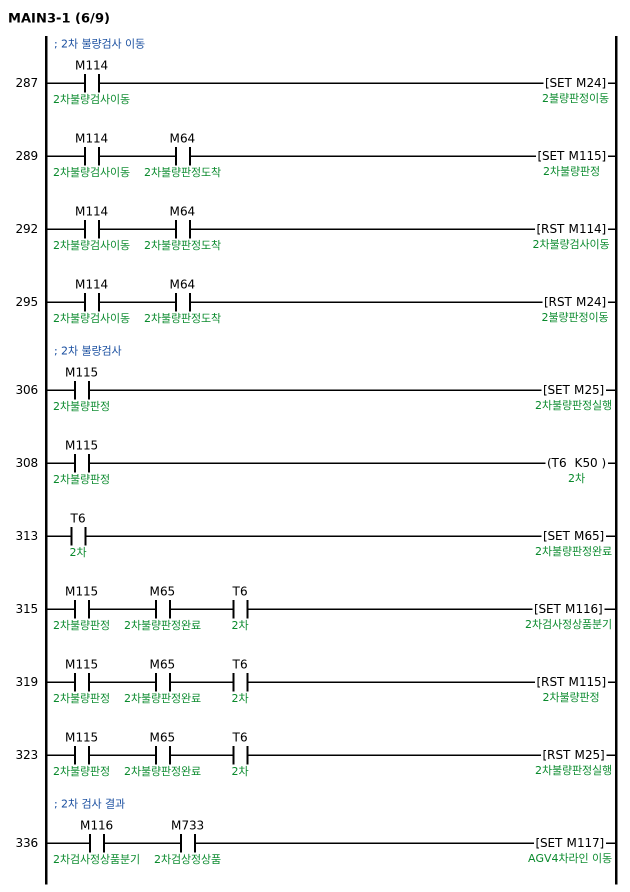
; 2차 불량검사 이동
287   LD      M114  ; 2차불량검사이동
      SET     M24  ; 2불량판정이동
289   LD      M114  ; 2차불량검사이동
      AND     M64  ; 2차불량판정도착
      SET     M115  ; 2차불량판정
292   LD      M114  ; 2차불량검사이동
      AND     M64  ; 2차불량판정도착
      RST     M114  ; 2차불량검사이동
295   LD      M114  ; 2차불량검사이동
      AND     M64  ; 2차불량판정도착
      RST     M24  ; 2불량판정이동
; 2차 불량검사
306   LD      M115  ; 2차불량판정
      SET     M25  ; 2차불량판정실행
308   LD      M115  ; 2차불량판정
      OUT     T6 K50  ; 2차
313   LD      T6  ; 2차
      SET     M65  ; 2차불량판정완료
315   LD      M115  ; 2차불량판정
      AND     M65  ; 2차불량판정완료
      AND     T6  ; 2차
      SET     M116  ; 2차검사정상품분기
319   LD      M115  ; 2차불량판정
      AND     M65  ; 2차불량판정완료
      AND     T6  ; 2차
      RST     M115  ; 2차불량판정
323   LD      M115  ; 2차불량판정
      AND     M65  ; 2차불량판정완료
      AND     T6  ; 2차
      RST     M25  ; 2차불량판정실행
; 2차 검사 결과
336   LD      M116  ; 2차검사정상품분기
      AND     M733  ; 2차검상정상품
      SET     M117  ; AGV4차라인 이동
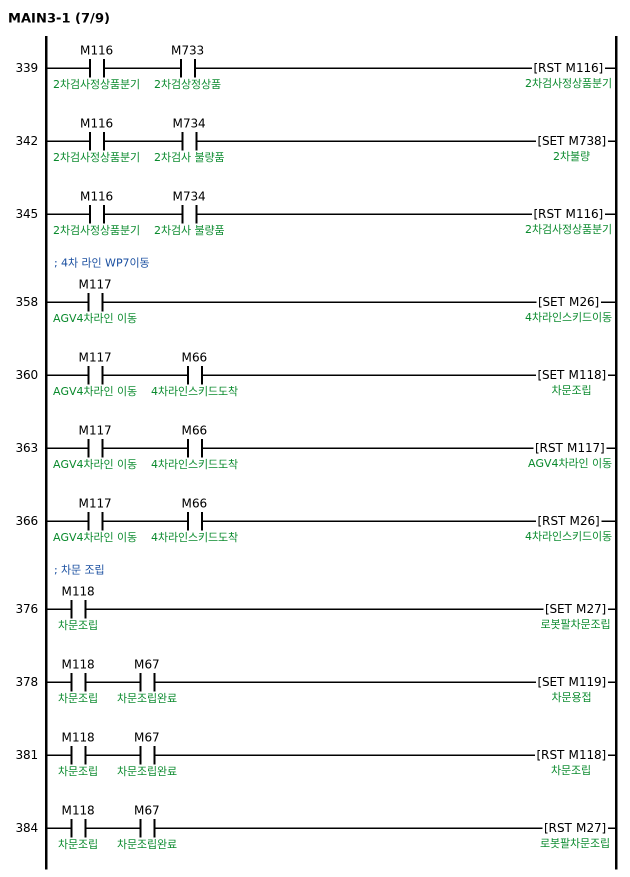
339   LD      M116  ; 2차검사정상품분기
      AND     M733  ; 2차검상정상품
      RST     M116  ; 2차검사정상품분기
342   LD      M116  ; 2차검사정상품분기
      AND     M734  ; 2차검사 불량품
      SET     M738  ; 2차불량
345   LD      M116  ; 2차검사정상품분기
      AND     M734  ; 2차검사 불량품
      RST     M116  ; 2차검사정상품분기
; 4차 라인 WP7이동
358   LD      M117  ; AGV4차라인 이동
      SET     M26  ; 4차라인스키드이동
360   LD      M117  ; AGV4차라인 이동
      AND     M66  ; 4차라인스키드도착
      SET     M118  ; 차문조립
363   LD      M117  ; AGV4차라인 이동
      AND     M66  ; 4차라인스키드도착
      RST     M117  ; AGV4차라인 이동
366   LD      M117  ; AGV4차라인 이동
      AND     M66  ; 4차라인스키드도착
      RST     M26  ; 4차라인스키드이동
; 차문 조립
376   LD      M118  ; 차문조립
      SET     M27  ; 로봇팔차문조립
378   LD      M118  ; 차문조립
      AND     M67  ; 차문조립완료
      SET     M119  ; 차문용접
381   LD      M118  ; 차문조립
      AND     M67  ; 차문조립완료
      RST     M118  ; 차문조립
384   LD      M118  ; 차문조립
      AND     M67  ; 차문조립완료
      RST     M27  ; 로봇팔차문조립
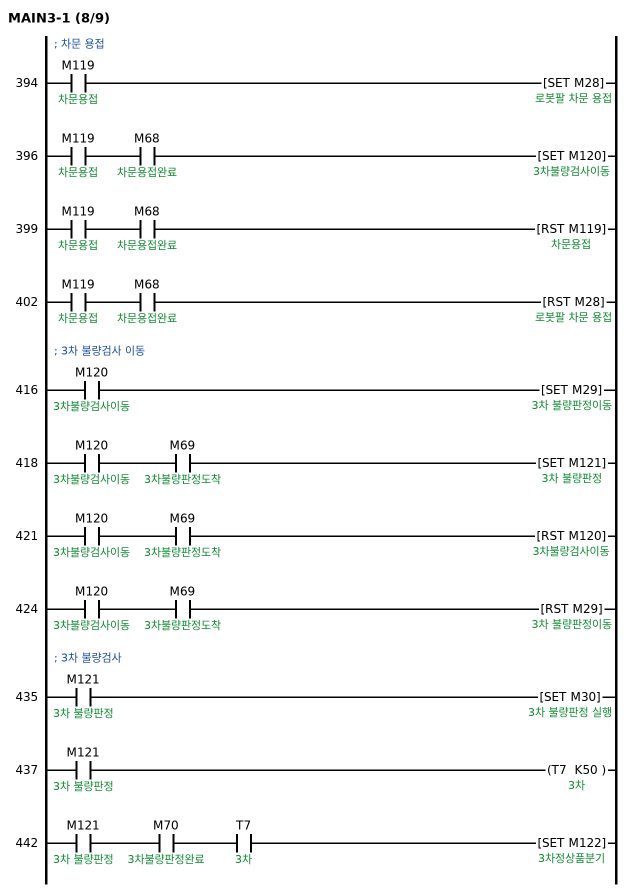
; 차문 용접
394   LD      M119  ; 차문용접
      SET     M28  ; 로봇팔 차문 용접
396   LD      M119  ; 차문용접
      AND     M68  ; 차문용접완료
      SET     M120  ; 3차불량검사이동
399   LD      M119  ; 차문용접
      AND     M68  ; 차문용접완료
      RST     M119  ; 차문용접
402   LD      M119  ; 차문용접
      AND     M68  ; 차문용접완료
      RST     M28  ; 로봇팔 차문 용접
; 3차 불량검사 이동
416   LD      M120  ; 3차불량검사이동
      SET     M29  ; 3차 불량판정이동
418   LD      M120  ; 3차불량검사이동
      AND     M69  ; 3차불량판정도착
      SET     M121  ; 3차 불량판정
421   LD      M120  ; 3차불량검사이동
      AND     M69  ; 3차불량판정도착
      RST     M120  ; 3차불량검사이동
424   LD      M120  ; 3차불량검사이동
      AND     M69  ; 3차불량판정도착
      RST     M29  ; 3차 불량판정이동
; 3차 불량검사
435   LD      M121  ; 3차 불량판정
      SET     M30  ; 3차 불량판정 실행
437   LD      M121  ; 3차 불량판정
      OUT     T7 K50  ; 3차
442   LD      M121  ; 3차 불량판정
      AND     M70  ; 3차불량판정완료
      AND     T7  ; 3차
      SET     M122  ; 3차정상품분기
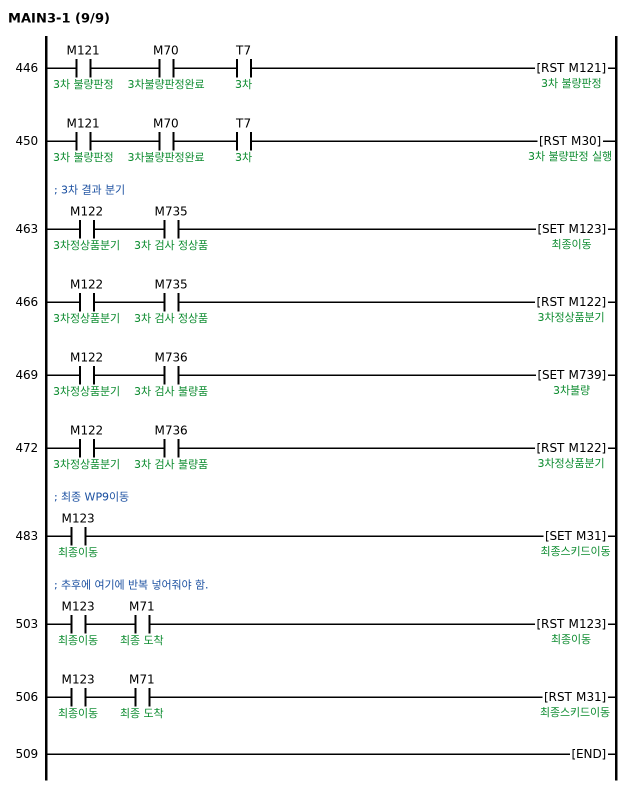
446   LD      M121  ; 3차 불량판정
      AND     M70  ; 3차불량판정완료
      AND     T7  ; 3차
      RST     M121  ; 3차 불량판정
450   LD      M121  ; 3차 불량판정
      AND     M70  ; 3차불량판정완료
      AND     T7  ; 3차
      RST     M30  ; 3차 불량판정 실행
; 3차 결과 분기
463   LD      M122  ; 3차정상품분기
      AND     M735  ; 3차 검사 정상품
      SET     M123  ; 최종이동
466   LD      M122  ; 3차정상품분기
      AND     M735  ; 3차 검사 정상품
      RST     M122  ; 3차정상품분기
469   LD      M122  ; 3차정상품분기
      AND     M736  ; 3차 검사 불량품
      SET     M739  ; 3차불량
472   LD      M122  ; 3차정상품분기
      AND     M736  ; 3차 검사 불량품
      RST     M122  ; 3차정상품분기
; 최종 WP9이동
483   LD      M123  ; 최종이동
      SET     M31  ; 최종스키드이동
; 추후에 여기에 반복 넣어줘야 함.
503   LD      M123  ; 최종이동
      AND     M71  ; 최종 도착
      RST     M123  ; 최종이동
506   LD      M123  ; 최종이동
      AND     M71  ; 최종 도착
      RST     M31  ; 최종스키드이동
509   END
END_PROGRAM

PROGRAM MAIN2-1
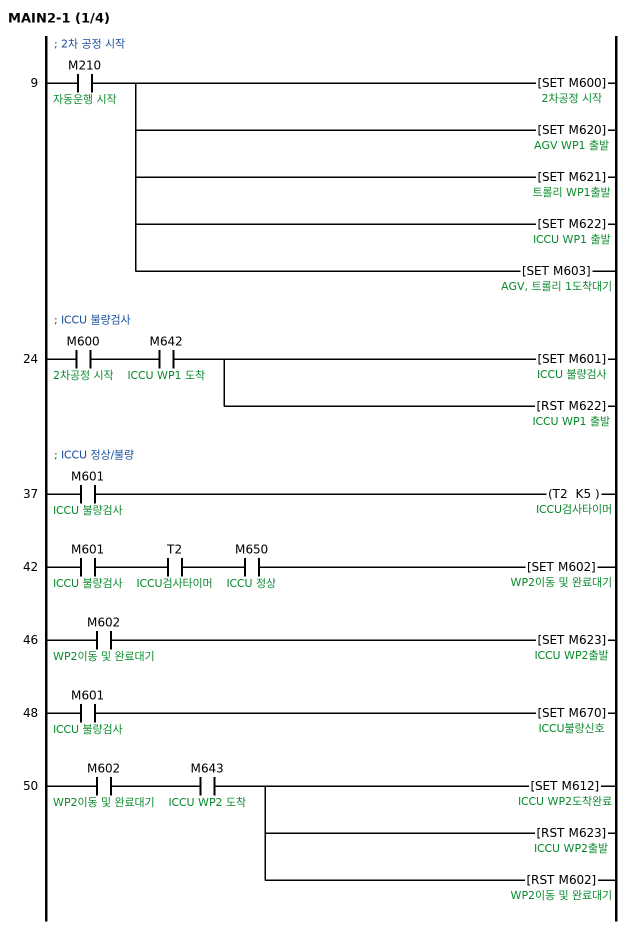
; 2차 공정 시작
9     LD      M210  ; 자동운행 시작
      SET     M600  ; 2차공정 시작
      SET     M620  ; AGV WP1 출발
      SET     M621  ; 트롤리 WP1출발
      SET     M622  ; ICCU WP1 출발
      SET     M603  ; AGV, 트롤리 1도착대기
; ICCU 불량검사
24    LD      M600  ; 2차공정 시작
      AND     M642  ; ICCU WP1 도착
      SET     M601  ; ICCU 불량검사
      RST     M622  ; ICCU WP1 출발
; ICCU 정상/불량
37    LD      M601  ; ICCU 불량검사
      OUT     T2 K5  ; ICCU검사타이머
42    LD      M601  ; ICCU 불량검사
      AND     T2  ; ICCU검사타이머
      AND     M650  ; ICCU 정상
      SET     M602  ; WP2이동 및 완료대기
46    LD      M602  ; WP2이동 및 완료대기
      SET     M623  ; ICCU WP2출발
48    LD      M601  ; ICCU 불량검사
      SET     M670  ; ICCU불량신호
50    LD      M602  ; WP2이동 및 완료대기
      AND     M643  ; ICCU WP2 도착
      SET     M612  ; ICCU WP2도착완료
      RST     M623  ; ICCU WP2출발
      RST     M602  ; WP2이동 및 완료대기
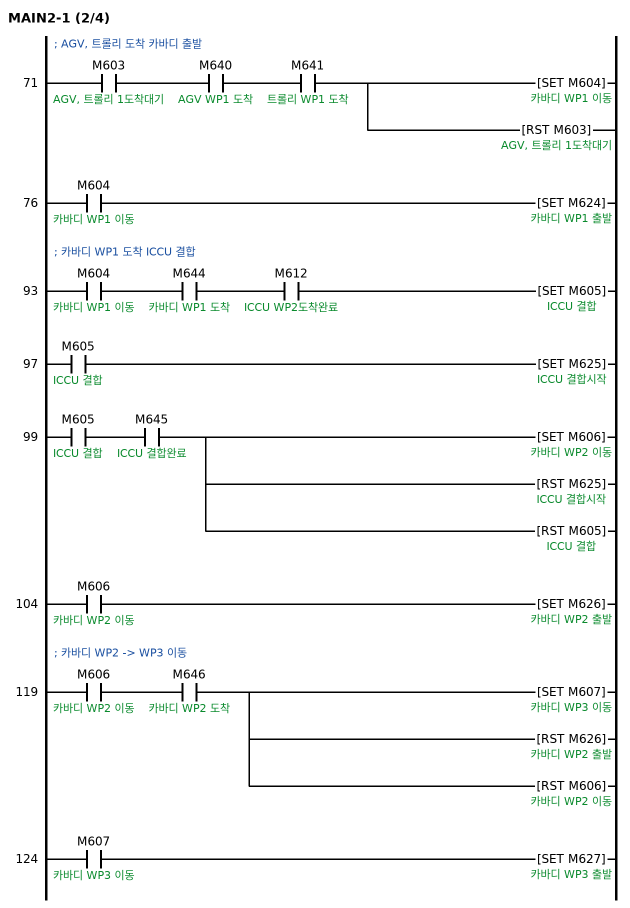
; AGV, 트롤리 도착 카바디 출발
71    LD      M603  ; AGV, 트롤리 1도착대기
      AND     M640  ; AGV WP1 도착
      AND     M641  ; 트롤리 WP1 도착
      SET     M604  ; 카바디 WP1 이동
      RST     M603  ; AGV, 트롤리 1도착대기
76    LD      M604  ; 카바디 WP1 이동
      SET     M624  ; 카바디 WP1 출발
; 카바디 WP1 도착 ICCU 결합
93    LD      M604  ; 카바디 WP1 이동
      AND     M644  ; 카바디 WP1 도착
      AND     M612  ; ICCU WP2도착완료
      SET     M605  ; ICCU 결합
97    LD      M605  ; ICCU 결합
      SET     M625  ; ICCU 결합시작
99    LD      M605  ; ICCU 결합
      AND     M645  ; ICCU 결합완료
      SET     M606  ; 카바디 WP2 이동
      RST     M625  ; ICCU 결합시작
      RST     M605  ; ICCU 결합
104   LD      M606  ; 카바디 WP2 이동
      SET     M626  ; 카바디 WP2 출발
; 카바디 WP2 -> WP3 이동
119   LD      M606  ; 카바디 WP2 이동
      AND     M646  ; 카바디 WP2 도착
      SET     M607  ; 카바디 WP3 이동
      RST     M626  ; 카바디 WP2 출발
      RST     M606  ; 카바디 WP2 이동
124   LD      M607  ; 카바디 WP3 이동
      SET     M627  ; 카바디 WP3 출발
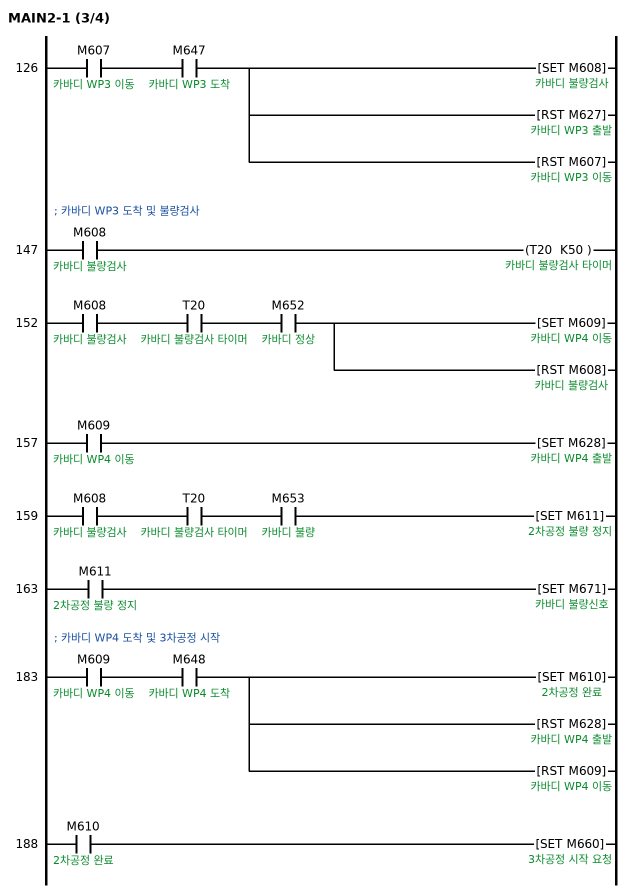
126   LD      M607  ; 카바디 WP3 이동
      AND     M647  ; 카바디 WP3 도착
      SET     M608  ; 카바디 불량검사
      RST     M627  ; 카바디 WP3 출발
      RST     M607  ; 카바디 WP3 이동
; 카바디 WP3 도착 및 불량검사
147   LD      M608  ; 카바디 불량검사
      OUT     T20 K50  ; 카바디 불량검사 타이머
152   LD      M608  ; 카바디 불량검사
      AND     T20  ; 카바디 불량검사 타이머
      AND     M652  ; 카바디 정상
      SET     M609  ; 카바디 WP4 이동
      RST     M608  ; 카바디 불량검사
157   LD      M609  ; 카바디 WP4 이동
      SET     M628  ; 카바디 WP4 출발
159   LD      M608  ; 카바디 불량검사
      AND     T20  ; 카바디 불량검사 타이머
      AND     M653  ; 카바디 불량
      SET     M611  ; 2차공정 불량 정지
163   LD      M611  ; 2차공정 불량 정지
      SET     M671  ; 카바디 불량신호
; 카바디 WP4 도착 및 3차공정 시작
183   LD      M609  ; 카바디 WP4 이동
      AND     M648  ; 카바디 WP4 도착
      SET     M610  ; 2차공정 완료
      RST     M628  ; 카바디 WP4 출발
      RST     M609  ; 카바디 WP4 이동
188   LD      M610  ; 2차공정 완료
      SET     M660  ; 3차공정 시작 요청
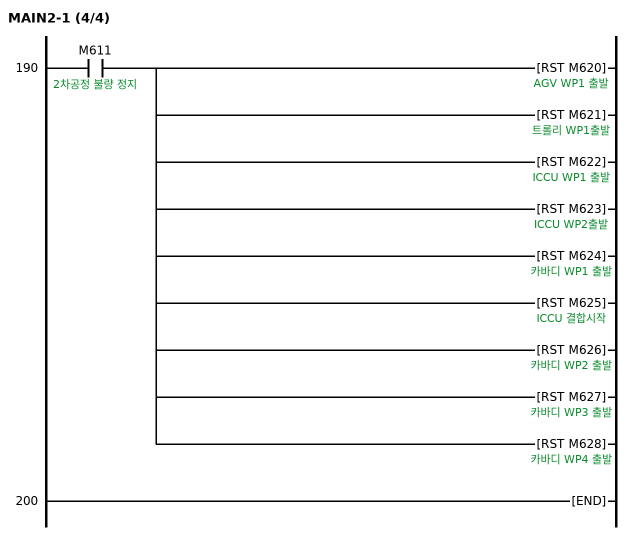
190   LD      M611  ; 2차공정 불량 정지
      RST     M620  ; AGV WP1 출발
      RST     M621  ; 트롤리 WP1출발
      RST     M622  ; ICCU WP1 출발
      RST     M623  ; ICCU WP2출발
      RST     M624  ; 카바디 WP1 출발
      RST     M625  ; ICCU 결합시작
      RST     M626  ; 카바디 WP2 출발
      RST     M627  ; 카바디 WP3 출발
      RST     M628  ; 카바디 WP4 출발
200   END
END_PROGRAM

PROGRAM MAIN2-2
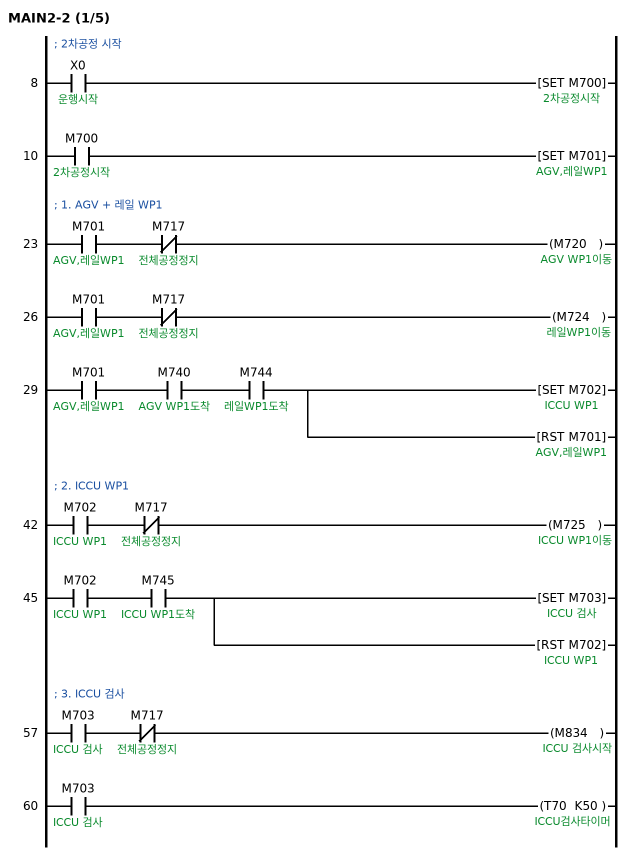
; 2차공정 시작
8     LD      X0  ; 운행시작
      SET     M700  ; 2차공정시작
10    LD      M700  ; 2차공정시작
      SET     M701  ; AGV,레일WP1
; 1. AGV + 레일 WP1
23    LD      M701  ; AGV,레일WP1
      ANI     M717  ; 전체공정정지
      OUT     M720  ; AGV WP1이동
26    LD      M701  ; AGV,레일WP1
      ANI     M717  ; 전체공정정지
      OUT     M724  ; 레일WP1이동
29    LD      M701  ; AGV,레일WP1
      AND     M740  ; AGV WP1도착
      AND     M744  ; 레일WP1도착
      SET     M702  ; ICCU WP1
      RST     M701  ; AGV,레일WP1
; 2. ICCU WP1
42    LD      M702  ; ICCU WP1
      ANI     M717  ; 전체공정정지
      OUT     M725  ; ICCU WP1이동
45    LD      M702  ; ICCU WP1
      AND     M745  ; ICCU WP1도착
      SET     M703  ; ICCU 검사
      RST     M702  ; ICCU WP1
; 3. ICCU 검사
57    LD      M703  ; ICCU 검사
      ANI     M717  ; 전체공정정지
      OUT     M834  ; ICCU 검사시작
60    LD      M703  ; ICCU 검사
      OUT     T70 K50  ; ICCU검사타이머
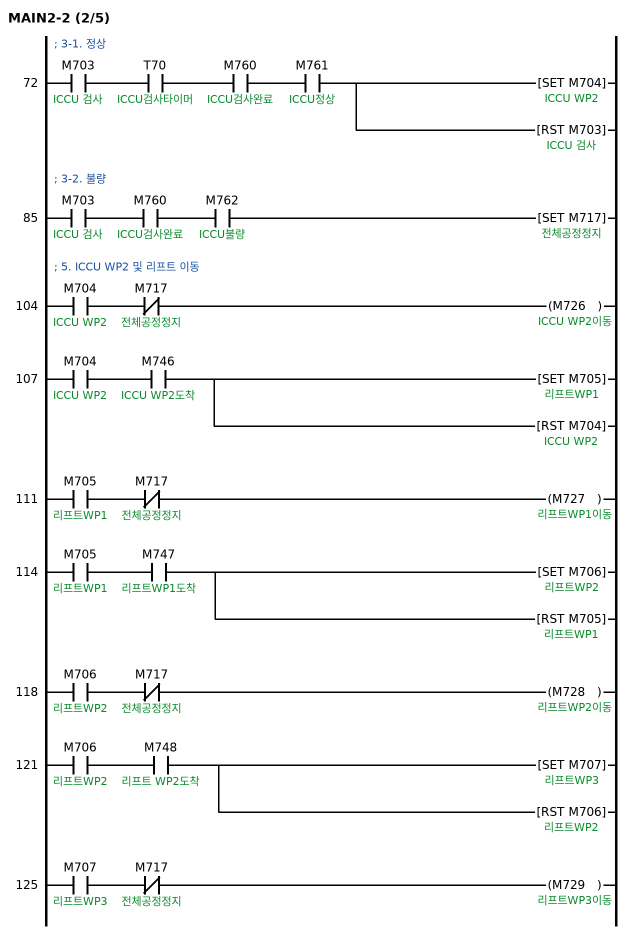
; 3-1. 정상
72    LD      M703  ; ICCU 검사
      AND     T70  ; ICCU검사타이머
      AND     M760  ; ICCU검사완료
      AND     M761  ; ICCU정상
      SET     M704  ; ICCU WP2
      RST     M703  ; ICCU 검사
; 3-2. 불량
85    LD      M703  ; ICCU 검사
      AND     M760  ; ICCU검사완료
      AND     M762  ; ICCU불량
      SET     M717  ; 전체공정정지
; 5. ICCU WP2 및 리프트 이동
104   LD      M704  ; ICCU WP2
      ANI     M717  ; 전체공정정지
      OUT     M726  ; ICCU WP2이동
107   LD      M704  ; ICCU WP2
      AND     M746  ; ICCU WP2도착
      SET     M705  ; 리프트WP1
      RST     M704  ; ICCU WP2
111   LD      M705  ; 리프트WP1
      ANI     M717  ; 전체공정정지
      OUT     M727  ; 리프트WP1이동
114   LD      M705  ; 리프트WP1
      AND     M747  ; 리프트WP1도착
      SET     M706  ; 리프트WP2
      RST     M705  ; 리프트WP1
118   LD      M706  ; 리프트WP2
      ANI     M717  ; 전체공정정지
      OUT     M728  ; 리프트WP2이동
121   LD      M706  ; 리프트WP2
      AND     M748  ; 리프트 WP2도착
      SET     M707  ; 리프트WP3
      RST     M706  ; 리프트WP2
125   LD      M707  ; 리프트WP3
      ANI     M717  ; 전체공정정지
      OUT     M729  ; 리프트WP3이동
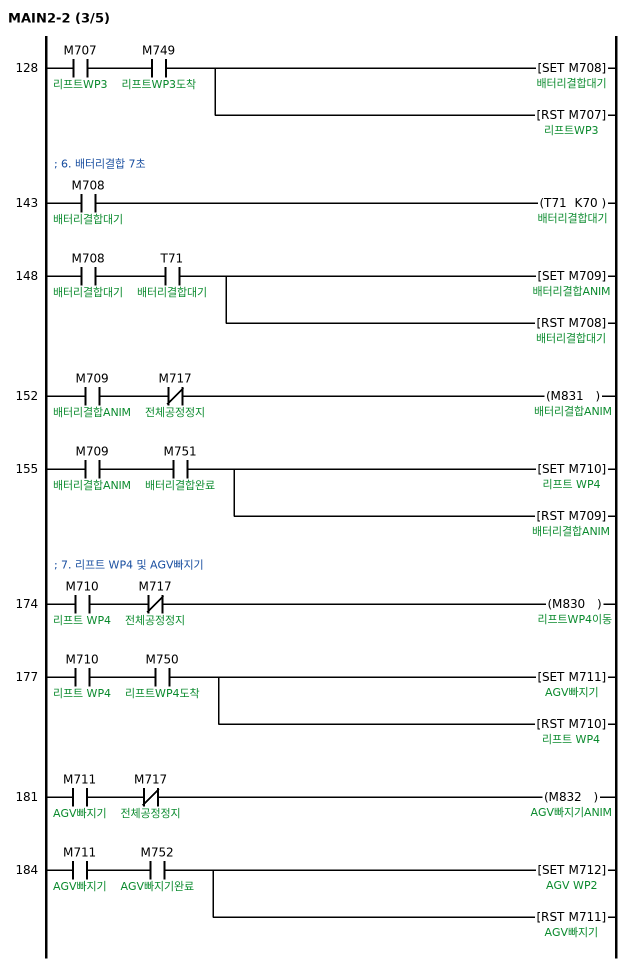
128   LD      M707  ; 리프트WP3
      AND     M749  ; 리프트WP3도착
      SET     M708  ; 배터리결합대기
      RST     M707  ; 리프트WP3
; 6. 배터리결합 7초
143   LD      M708  ; 배터리결합대기
      OUT     T71 K70  ; 배터리결합대기
148   LD      M708  ; 배터리결합대기
      AND     T71  ; 배터리결합대기
      SET     M709  ; 배터리결합ANIM
      RST     M708  ; 배터리결합대기
152   LD      M709  ; 배터리결합ANIM
      ANI     M717  ; 전체공정정지
      OUT     M831  ; 배터리결합ANIM
155   LD      M709  ; 배터리결합ANIM
      AND     M751  ; 배터리결합완료
      SET     M710  ; 리프트 WP4
      RST     M709  ; 배터리결합ANIM
; 7. 리프트 WP4 및 AGV빠지기
174   LD      M710  ; 리프트 WP4
      ANI     M717  ; 전체공정정지
      OUT     M830  ; 리프트WP4이동
177   LD      M710  ; 리프트 WP4
      AND     M750  ; 리프트WP4도착
      SET     M711  ; AGV빠지기
      RST     M710  ; 리프트 WP4
181   LD      M711  ; AGV빠지기
      ANI     M717  ; 전체공정정지
      OUT     M832  ; AGV빠지기ANIM
184   LD      M711  ; AGV빠지기
      AND     M752  ; AGV빠지기완료
      SET     M712  ; AGV WP2
      RST     M711  ; AGV빠지기
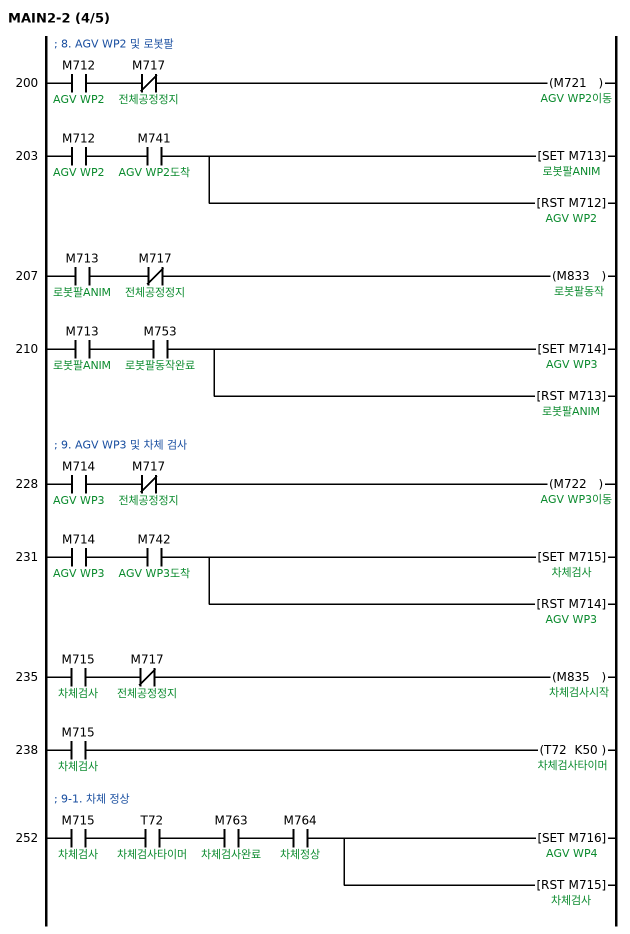
; 8. AGV WP2 및 로봇팔
200   LD      M712  ; AGV WP2
      ANI     M717  ; 전체공정정지
      OUT     M721  ; AGV WP2이동
203   LD      M712  ; AGV WP2
      AND     M741  ; AGV WP2도착
      SET     M713  ; 로봇팔ANIM
      RST     M712  ; AGV WP2
207   LD      M713  ; 로봇팔ANIM
      ANI     M717  ; 전체공정정지
      OUT     M833  ; 로봇팔동작
210   LD      M713  ; 로봇팔ANIM
      AND     M753  ; 로봇팔동작완료
      SET     M714  ; AGV WP3
      RST     M713  ; 로봇팔ANIM
; 9. AGV WP3 및 차체 검사
228   LD      M714  ; AGV WP3
      ANI     M717  ; 전체공정정지
      OUT     M722  ; AGV WP3이동
231   LD      M714  ; AGV WP3
      AND     M742  ; AGV WP3도착
      SET     M715  ; 차체검사
      RST     M714  ; AGV WP3
235   LD      M715  ; 차체검사
      ANI     M717  ; 전체공정정지
      OUT     M835  ; 차체검사시작
238   LD      M715  ; 차체검사
      OUT     T72 K50  ; 차체검사타이머
; 9-1. 차체 정상
252   LD      M715  ; 차체검사
      AND     T72  ; 차체검사타이머
      AND     M763  ; 차체검사완료
      AND     M764  ; 차체정상
      SET     M716  ; AGV WP4
      RST     M715  ; 차체검사
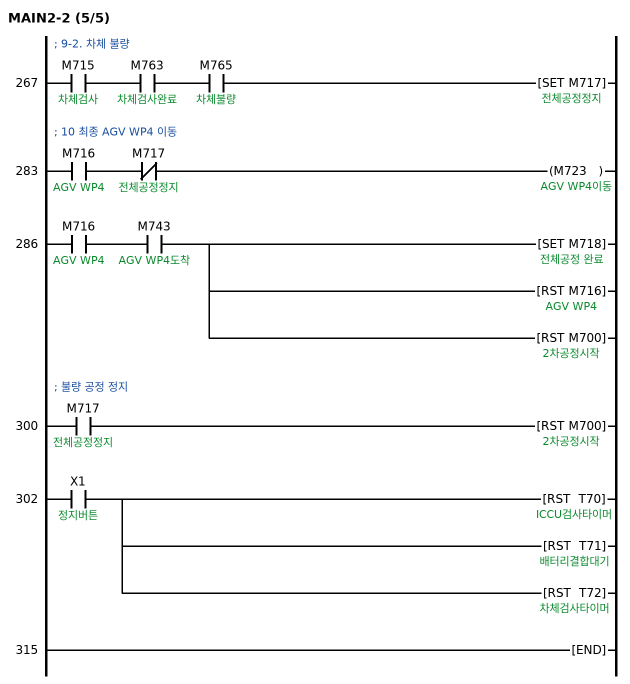
; 9-2. 차체 불량
267   LD      M715  ; 차체검사
      AND     M763  ; 차체검사완료
      AND     M765  ; 차체불량
      SET     M717  ; 전체공정정지
; 10 최종 AGV WP4 이동
283   LD      M716  ; AGV WP4
      ANI     M717  ; 전체공정정지
      OUT     M723  ; AGV WP4이동
286   LD      M716  ; AGV WP4
      AND     M743  ; AGV WP4도착
      SET     M718  ; 전체공정 완료
      RST     M716  ; AGV WP4
      RST     M700  ; 2차공정시작
; 불량 공정 정지
300   LD      M717  ; 전체공정정지
      RST     M700  ; 2차공정시작
302   LD      X1  ; 정지버튼
      RST     T70  ; ICCU검사타이머
      RST     T71  ; 배터리결합대기
      RST     T72  ; 차체검사타이머
315   END
END_PROGRAM

PROGRAM MAIN3-T
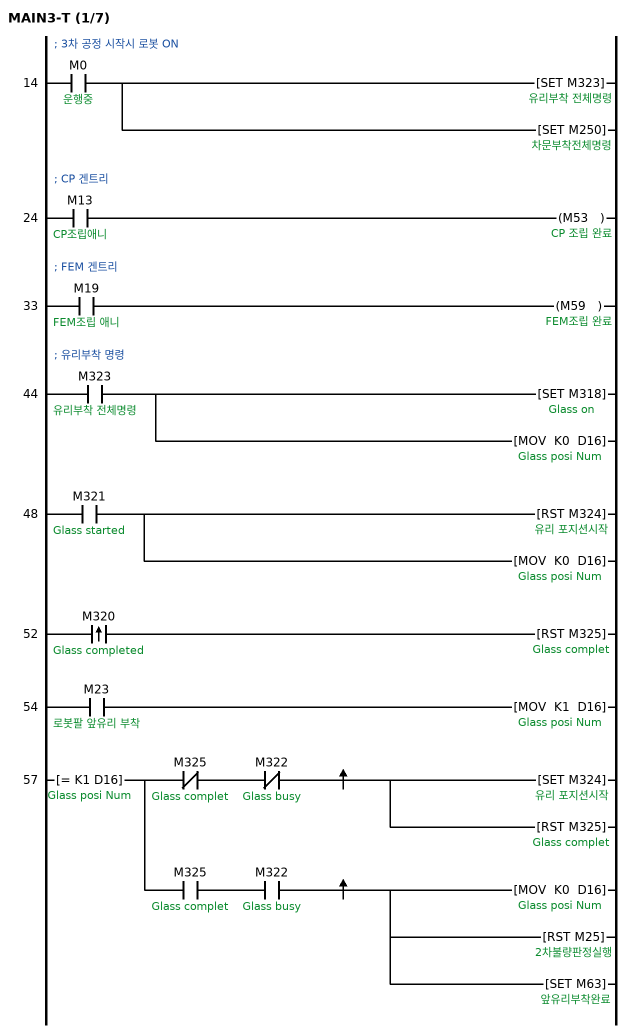
; 3차 공정 시작시 로봇 ON
14    LD      M0  ; 운행중
      SET     M323  ; 유리부착 전체명령
      SET     M250  ; 차문부착전체명령
; CP 겐트리
24    LD      M13  ; CP조립애니
      OUT     M53  ; CP 조립 완료
; FEM 겐트리
33    LD      M19  ; FEM조립 애니
      OUT     M59  ; FEM조립 완료
; 유리부착 명령
44    LD      M323  ; 유리부착 전체명령
      SET     M318  ; Glass on
      MOV     K0 D16  ; Glass posi Num
48    LD      M321  ; Glass started
      RST     M324  ; 유리 포지션시작
      MOV     K0 D16
52    LDP     M320  ; Glass completed
      RST     M325  ; Glass complet
54    LD      M23  ; 로봇팔 앞유리 부착
      MOV     K1 D16
57    LD=     K1 D16  ; Glass posi Num
      MPS
      ANI     M325  ; Glass complet
      ANI     M322  ; Glass busy
      MEP
      SET     M324  ; 유리 포지션시작
      RST     M325  ; Glass complet
      MPP
      AND     M325  ; Glass complet
      AND     M322  ; Glass busy
      MEP
      MOV     K0 D16
      RST     M25  ; 2차불량판정실행
      SET     M63  ; 앞유리부착완료
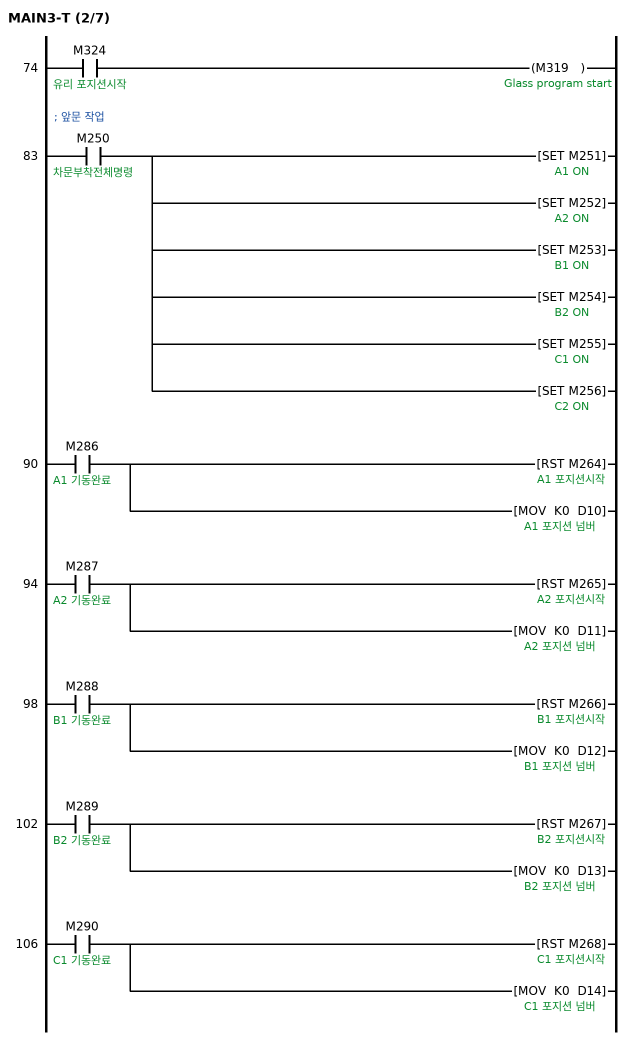
74    LD      M324  ; 유리 포지션시작
      OUT     M319  ; Glass program start
; 앞문 작업
83    LD      M250  ; 차문부착전체명령
      SET     M251  ; A1 ON
      SET     M252  ; A2 ON
      SET     M253  ; B1 ON
      SET     M254  ; B2 ON
      SET     M255  ; C1 ON
      SET     M256  ; C2 ON
90    LD      M286  ; A1 기동완료
      RST     M264  ; A1 포지션시작
      MOV     K0 D10  ; A1 포지션 넘버
94    LD      M287  ; A2 기동완료
      RST     M265  ; A2 포지션시작
      MOV     K0 D11  ; A2 포지션 넘버
98    LD      M288  ; B1 기동완료
      RST     M266  ; B1 포지션시작
      MOV     K0 D12  ; B1 포지션 넘버
102   LD      M289  ; B2 기동완료
      RST     M267  ; B2 포지션시작
      MOV     K0 D13  ; B2 포지션 넘버
106   LD      M290  ; C1 기동완료
      RST     M268  ; C1 포지션시작
      MOV     K0 D14  ; C1 포지션 넘버
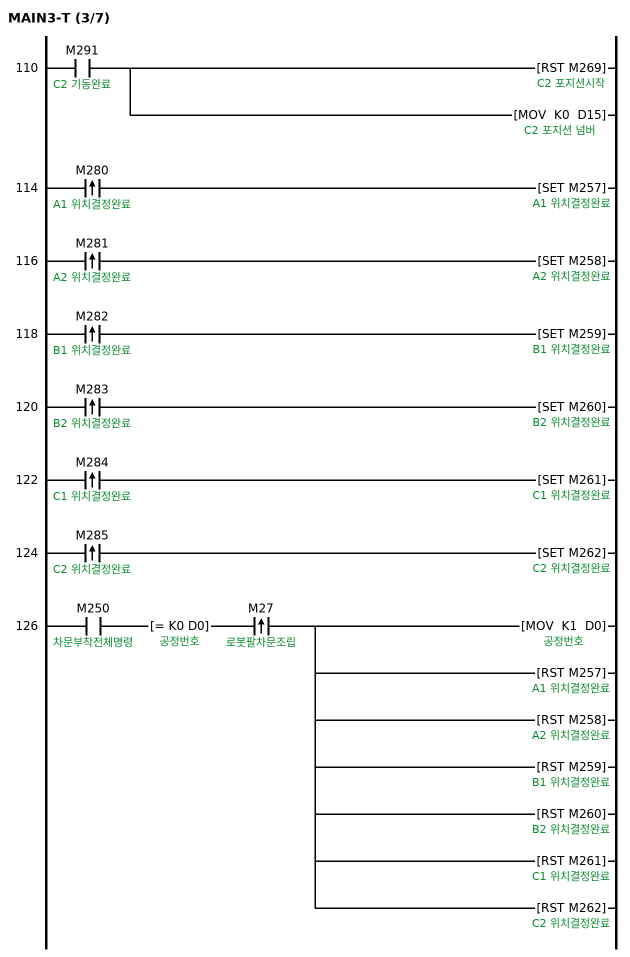
110   LD      M291  ; C2 기동완료
      RST     M269  ; C2 포지션시작
      MOV     K0 D15  ; C2 포지션 넘버
114   LDP     M280  ; A1 위치결정완료
      SET     M257  ; A1 위치결정완료
116   LDP     M281  ; A2 위치결정완료
      SET     M258  ; A2 위치결정완료
118   LDP     M282  ; B1 위치결정완료
      SET     M259  ; B1 위치결정완료
120   LDP     M283  ; B2 위치결정완료
      SET     M260  ; B2 위치결정완료
122   LDP     M284  ; C1 위치결정완료
      SET     M261  ; C1 위치결정완료
124   LDP     M285  ; C2 위치결정완료
      SET     M262  ; C2 위치결정완료
126   LD      M250  ; 차문부착전체명령
      AND=    K0 D0  ; 공정번호
      ANDP    M27  ; 로봇팔차문조립
      MOV     K1 D0
      RST     M257  ; A1 위치결정완료
      RST     M258  ; A2 위치결정완료
      RST     M259  ; B1 위치결정완료
      RST     M260  ; B2 위치결정완료
      RST     M261  ; C1 위치결정완료
      RST     M262  ; C2 위치결정완료
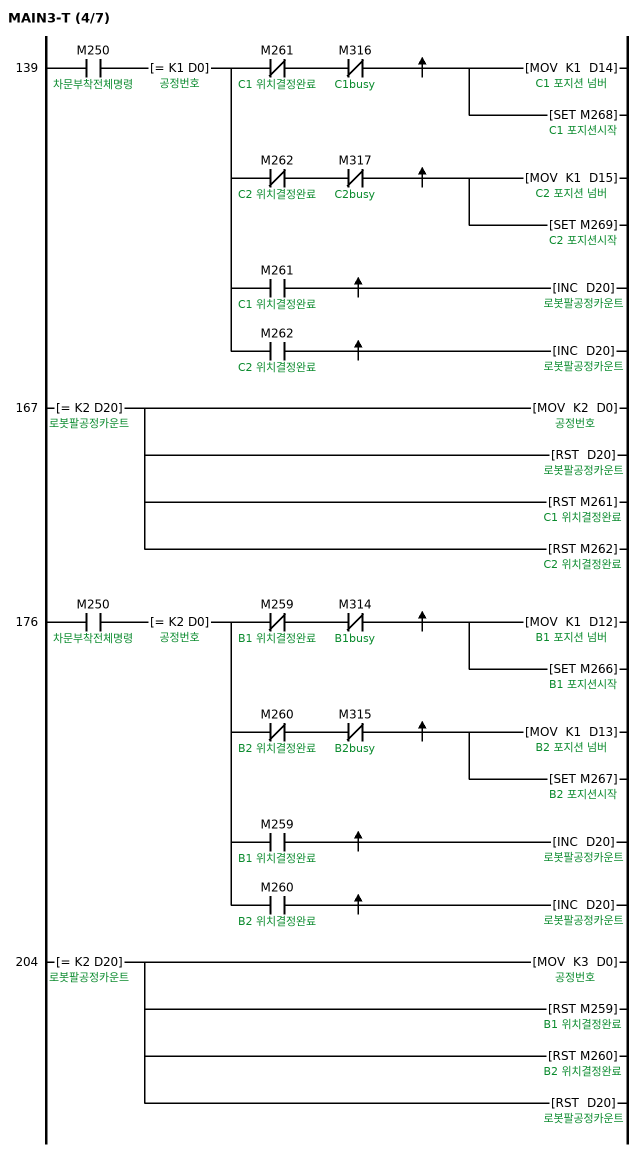
139   LD      M250  ; 차문부착전체명령
      AND=    K1 D0  ; 공정번호
      MPS
      ANI     M261  ; C1 위치결정완료
      ANI     M316  ; C1busy
      MEP
      MOV     K1 D14
      SET     M268  ; C1 포지션시작
      MRD
      ANI     M262  ; C2 위치결정완료
      ANI     M317  ; C2busy
      MEP
      MOV     K1 D15
      SET     M269  ; C2 포지션시작
      MRD
      AND     M261  ; C1 위치결정완료
      MEP
      INC     D20  ; 로봇팔공정카운트
      MPP
      AND     M262  ; C2 위치결정완료
      MEP
      INC     D20
167   LD=     K2 D20  ; 로봇팔공정카운트
      MOV     K2 D0
      RST     D20  ; 로봇팔공정카운트
      RST     M261  ; C1 위치결정완료
      RST     M262  ; C2 위치결정완료
176   LD      M250  ; 차문부착전체명령
      AND=    K2 D0  ; 공정번호
      MPS
      ANI     M259  ; B1 위치결정완료
      ANI     M314  ; B1busy
      MEP
      MOV     K1 D12
      SET     M266  ; B1 포지션시작
      MRD
      ANI     M260  ; B2 위치결정완료
      ANI     M315  ; B2busy
      MEP
      MOV     K1 D13
      SET     M267  ; B2 포지션시작
      MRD
      AND     M259  ; B1 위치결정완료
      MEP
      INC     D20
      MPP
      AND     M260  ; B2 위치결정완료
      MEP
      INC     D20
204   LD=     K2 D20  ; 로봇팔공정카운트
      MOV     K3 D0
      RST     M259  ; B1 위치결정완료
      RST     M260  ; B2 위치결정완료
      RST     D20  ; 로봇팔공정카운트
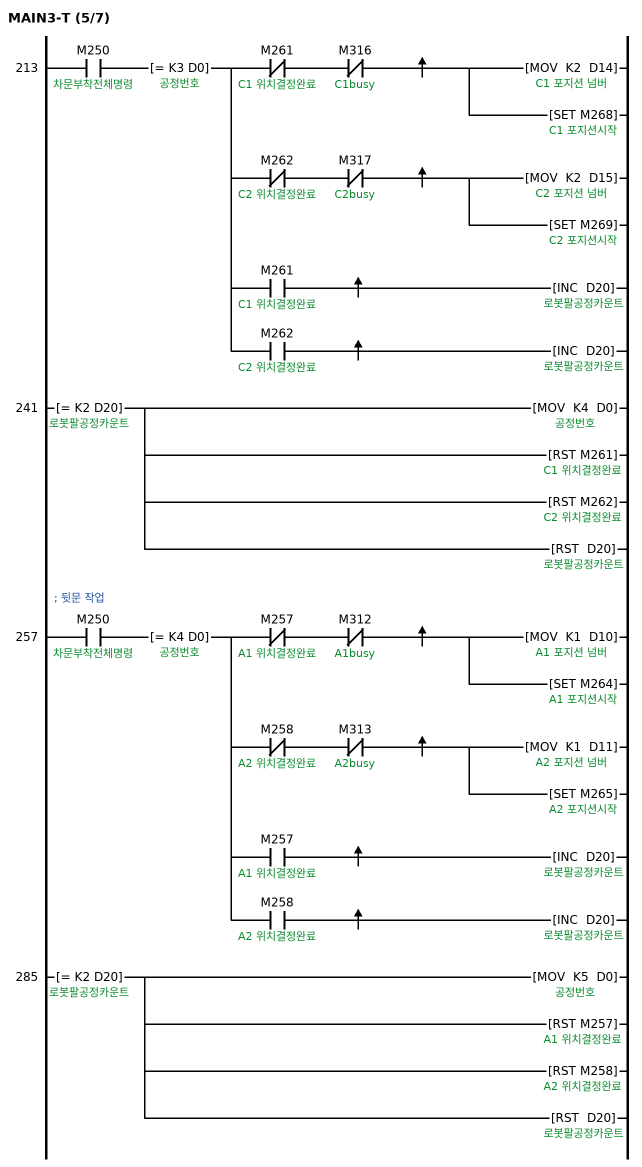
213   LD      M250  ; 차문부착전체명령
      AND=    K3 D0  ; 공정번호
      MPS
      ANI     M261  ; C1 위치결정완료
      ANI     M316  ; C1busy
      MEP
      MOV     K2 D14
      SET     M268  ; C1 포지션시작
      MRD
      ANI     M262  ; C2 위치결정완료
      ANI     M317  ; C2busy
      MEP
      MOV     K2 D15
      SET     M269  ; C2 포지션시작
      MRD
      AND     M261  ; C1 위치결정완료
      MEP
      INC     D20
      MPP
      AND     M262  ; C2 위치결정완료
      MEP
      INC     D20
241   LD=     K2 D20  ; 로봇팔공정카운트
      MOV     K4 D0
      RST     M261  ; C1 위치결정완료
      RST     M262  ; C2 위치결정완료
      RST     D20  ; 로봇팔공정카운트
; 뒷문 작업
257   LD      M250  ; 차문부착전체명령
      AND=    K4 D0  ; 공정번호
      MPS
      ANI     M257  ; A1 위치결정완료
      ANI     M312  ; A1busy
      MEP
      MOV     K1 D10
      SET     M264  ; A1 포지션시작
      MRD
      ANI     M258  ; A2 위치결정완료
      ANI     M313  ; A2busy
      MEP
      MOV     K1 D11
      SET     M265  ; A2 포지션시작
      MRD
      AND     M257  ; A1 위치결정완료
      MEP
      INC     D20
      MPP
      AND     M258  ; A2 위치결정완료
      MEP
      INC     D20
285   LD=     K2 D20  ; 로봇팔공정카운트
      MOV     K5 D0
      RST     M257  ; A1 위치결정완료
      RST     M258  ; A2 위치결정완료
      RST     D20  ; 로봇팔공정카운트
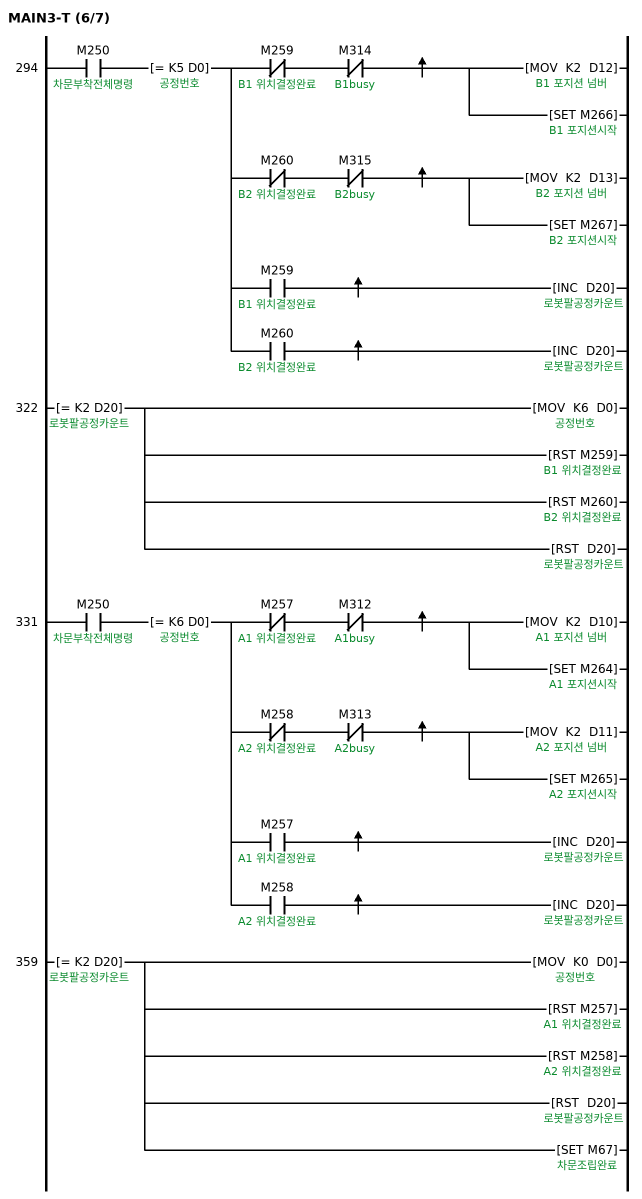
294   LD      M250  ; 차문부착전체명령
      AND=    K5 D0  ; 공정번호
      MPS
      ANI     M259  ; B1 위치결정완료
      ANI     M314  ; B1busy
      MEP
      MOV     K2 D12
      SET     M266  ; B1 포지션시작
      MRD
      ANI     M260  ; B2 위치결정완료
      ANI     M315  ; B2busy
      MEP
      MOV     K2 D13
      SET     M267  ; B2 포지션시작
      MRD
      AND     M259  ; B1 위치결정완료
      MEP
      INC     D20
      MPP
      AND     M260  ; B2 위치결정완료
      MEP
      INC     D20
322   LD=     K2 D20  ; 로봇팔공정카운트
      MOV     K6 D0
      RST     M259  ; B1 위치결정완료
      RST     M260  ; B2 위치결정완료
      RST     D20  ; 로봇팔공정카운트
331   LD      M250  ; 차문부착전체명령
      AND=    K6 D0  ; 공정번호
      MPS
      ANI     M257  ; A1 위치결정완료
      ANI     M312  ; A1busy
      MEP
      MOV     K2 D10
      SET     M264  ; A1 포지션시작
      MRD
      ANI     M258  ; A2 위치결정완료
      ANI     M313  ; A2busy
      MEP
      MOV     K2 D11
      SET     M265  ; A2 포지션시작
      MRD
      AND     M257  ; A1 위치결정완료
      MEP
      INC     D20
      MPP
      AND     M258  ; A2 위치결정완료
      MEP
      INC     D20
359   LD=     K2 D20  ; 로봇팔공정카운트
      MOV     K0 D0
      RST     M257  ; A1 위치결정완료
      RST     M258  ; A2 위치결정완료
      RST     D20  ; 로봇팔공정카운트
      SET     M67  ; 차문조립완료
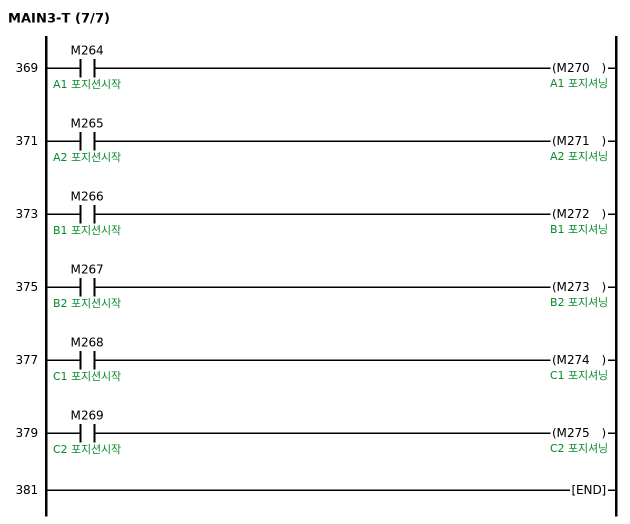
369   LD      M264  ; A1 포지션시작
      OUT     M270  ; A1 포지셔닝
371   LD      M265  ; A2 포지션시작
      OUT     M271  ; A2 포지셔닝
373   LD      M266  ; B1 포지션시작
      OUT     M272  ; B1 포지셔닝
375   LD      M267  ; B2 포지션시작
      OUT     M273  ; B2 포지셔닝
377   LD      M268  ; C1 포지션시작
      OUT     M274  ; C1 포지셔닝
379   LD      M269  ; C2 포지션시작
      OUT     M275  ; C2 포지셔닝
381   END
END_PROGRAM

// device comments not shown above
M32  ; 겐트리1 이동시작
M33  ; CP 조립 ANIM 시작
M34  ; 3-1불량판정시작
M40  ; 겐트리2 이동시작
M41  ; FEM 이동 시작
M42  ; 겐트리 이동 완료
M43  ; CP조립완료
M44  ; 3-1불량이동완료
M150  ; 1-1차전진완료
M151  ; 1-1불량판정완료
M152  ; 1-2레일전진완료
M153  ; AGV1차라인도착
M154  ; 커버조립 완료
M155  ; AGV2차라인 도착
M156  ; 1-2불량판정완료
M157  ; AGV2차공정도착
M200  ; 자동운행 시작
M201  ; AGV1차전진
M202  ; 커버1차전진
M203  ; 1-1불량판정 실행
M204  ; 커버레일2차전진
M205  ; 배터리팩커버조립
M206  ; AGV2차 라인 이동
M207  ; 1-2불량판정실행
M230  ; AGV+차체1이동
M231  ; 배터리결합
M232  ; ICCU 1 이동
M233  ; ICCU 불량검사 시작
M234  ; ICCU 2 이동
M235  ; ICCU 결합
M236  ; 차체 2 이동
M237  ; 차체 3 이동
M238  ; 차체 불량검사 시작
M239  ; 차체 4 이동
M240  ; 2번공정완료
M248  ; 유리 부착 프로그램 실행
M295  ; 차문 전체 완료
M326  ; Glass start
M330  ; C1 전원ON
M401  ; 1-1차불량판정
M402  ; 1-2라인이동,커버조립
M403  ; 1-2차 불량판정
M404  ; 1-2공정이동
M410  ; 1-1차레일전진
M411  ; 3-1불량판정
M412  ; 공정 3단계
M413  ; 공정 4단계
M414  ; 공정 5단계
M415  ; 공정 6단계
M416  ; 공정 7단계
M532  ; 1차 판정 유효
M535  ; 2차 판정결과 유효
M613  ; ICCU 결합 완료
M614  ; 롤러 차체 이동
M615  ; 차체 2 도착
M616  ; 차체 3 이동
M617  ; 차체 3 도착
M618  ; 차체 4 이동
M619  ; 차체 정상
C0  ; 3-1불량판정 카운트
C10  ; 로봇팔공정카운트
T10  ; ICCU검사타이머
T11  ; 차체 불량검사 타이머
T100  ; 앞유리  대기
